Fanuc KAREL source: kt00537.KL

-- PROVISIONAL review KL for V770-1; original PC SHA256 ffb0772971f6a8f15e09168681dae37f0a47dae6e722e0d7e489b6582cb7a491
-- Incomplete behavior may be omitted. Consult companion uncertainty JSON. Do not deploy.
PROGRAM KT00537
%NOLOCKGROUP
-- UNRESOLVED_DECL P1 type=000199
-- UNRESOLVED_DECL P2 type=000101
-- UNRESOLVED_DECL OUT type=000199
BEGIN
  -- UNRESOLVED_PC offsets 5-39; opcodes 49,7E,49,60,7E,4A
  -- UNRESOLVED_PC offsets 44-48; opcodes 7F
END KT00537
